// Mitsubishi GX Works2 project: PCL_레더   PLC: Q02/Q02H

PROGRAM MAIN
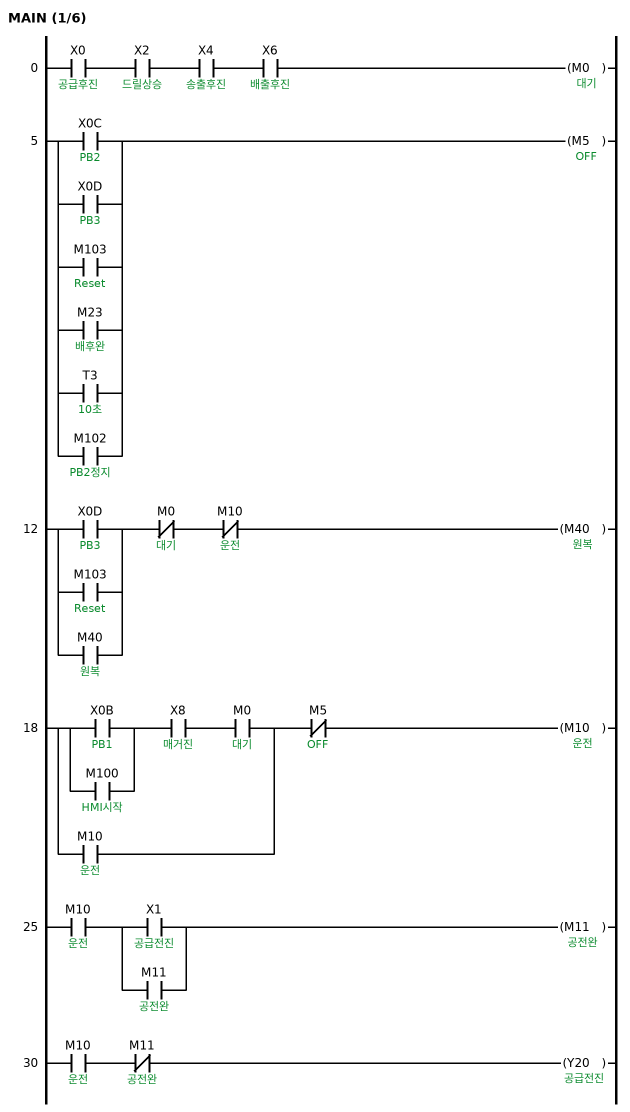
0     LD      X0  ; 공급후진
      AND     X2  ; 드릴상승
      AND     X4  ; 송출후진
      AND     X6  ; 배출후진
      OUT     M0  ; 대기
5     LD      X0C  ; PB2
      OR      X0D  ; PB3
      OR      M103  ; Reset
      OR      M23  ; 배후완
      OR      T3  ; 10초
      OR      M102  ; PB2정지
      OUT     M5  ; OFF
12    LD      X0D  ; PB3
      OR      M103  ; Reset
      OR      M40  ; 원복
      ANI     M0  ; 대기
      ANI     M10  ; 운전
      OUT     M40  ; 원복
18    LD      X0B  ; PB1
      OR      M100  ; HMI시작
      AND     X8  ; 매거진
      AND     M0  ; 대기
      OR      M10  ; 운전
      ANI     M5  ; OFF
      OUT     M10  ; 운전
25    LD      M10  ; 운전
      LD      X1  ; 공급전진
      OR      M11  ; 공전완
      ANB
      OUT     M11  ; 공전완
30    LD      M10  ; 운전
      ANI     M11  ; 공전완
      OUT     Y20  ; 공급전진
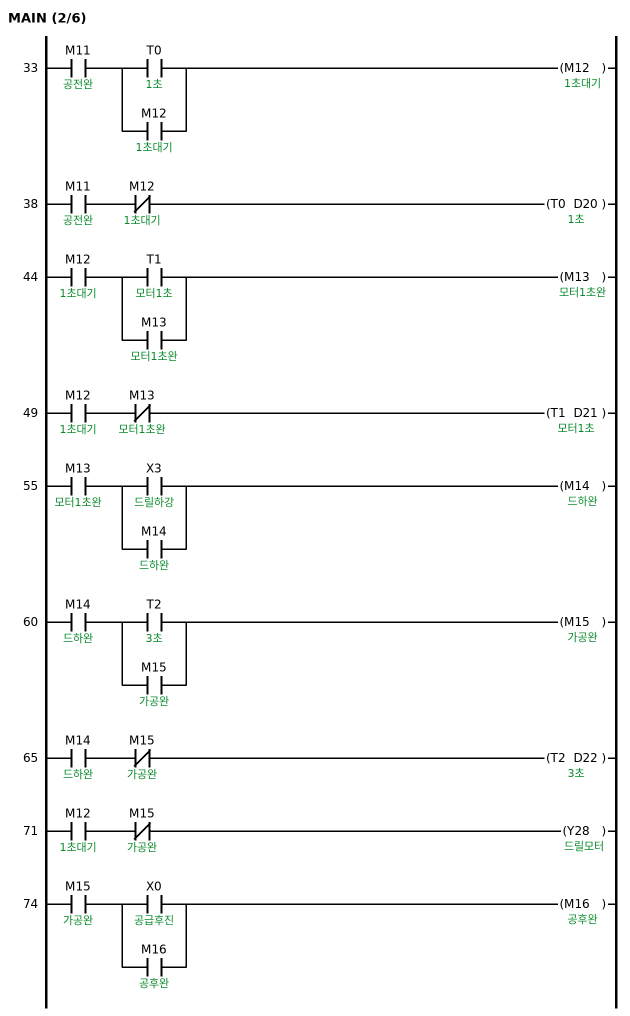
33    LD      M11  ; 공전완
      LD      T0  ; 1초
      OR      M12  ; 1초대기
      ANB
      OUT     M12  ; 1초대기
38    LD      M11  ; 공전완
      ANI     M12  ; 1초대기
      OUT     T0 D20  ; 1초
44    LD      M12  ; 1초대기
      LD      T1  ; 모터1초
      OR      M13  ; 모터1초완
      ANB
      OUT     M13  ; 모터1초완
49    LD      M12  ; 1초대기
      ANI     M13  ; 모터1초완
      OUT     T1 D21  ; 모터1초
55    LD      M13  ; 모터1초완
      LD      X3  ; 드릴하강
      OR      M14  ; 드하완
      ANB
      OUT     M14  ; 드하완
60    LD      M14  ; 드하완
      LD      T2  ; 3초
      OR      M15  ; 가공완
      ANB
      OUT     M15  ; 가공완
65    LD      M14  ; 드하완
      ANI     M15  ; 가공완
      OUT     T2 D22  ; 3초
71    LD      M12  ; 1초대기
      ANI     M15  ; 가공완
      OUT     Y28  ; 드릴모터
74    LD      M15  ; 가공완
      LD      X0  ; 공급후진
      OR      M16  ; 공후완
      ANB
      OUT     M16  ; 공후완
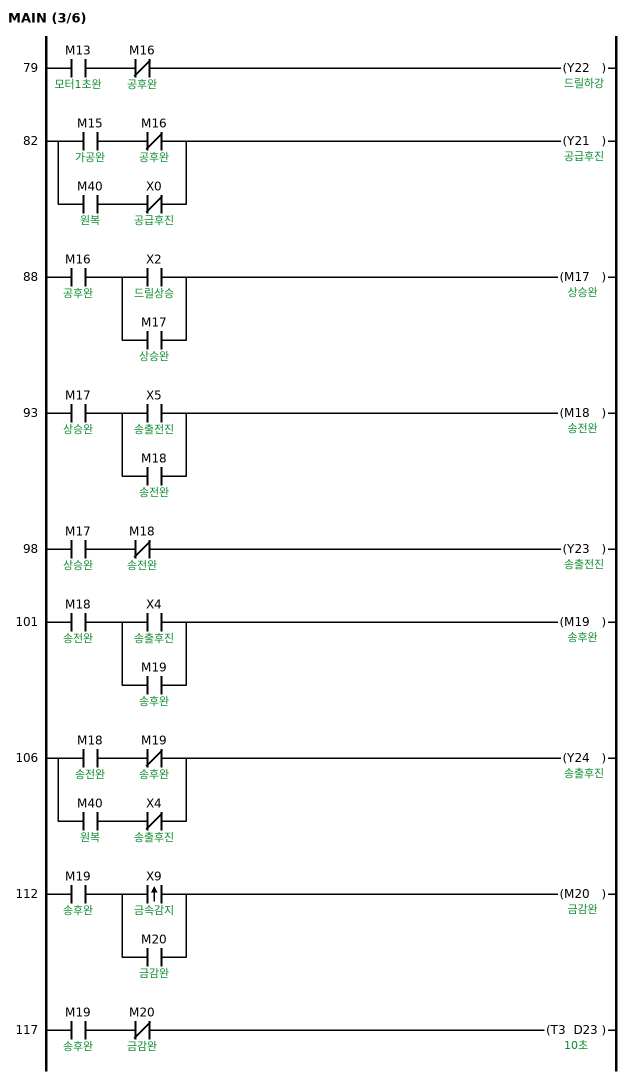
79    LD      M13  ; 모터1초완
      ANI     M16  ; 공후완
      OUT     Y22  ; 드릴하강
82    LD      M15  ; 가공완
      ANI     M16  ; 공후완
      LD      M40  ; 원복
      ANI     X0  ; 공급후진
      ORB
      OUT     Y21  ; 공급후진
88    LD      M16  ; 공후완
      LD      X2  ; 드릴상승
      OR      M17  ; 상승완
      ANB
      OUT     M17  ; 상승완
93    LD      M17  ; 상승완
      LD      X5  ; 송출전진
      OR      M18  ; 송전완
      ANB
      OUT     M18  ; 송전완
98    LD      M17  ; 상승완
      ANI     M18  ; 송전완
      OUT     Y23  ; 송출전진
101   LD      M18  ; 송전완
      LD      X4  ; 송출후진
      OR      M19  ; 송후완
      ANB
      OUT     M19  ; 송후완
106   LD      M18  ; 송전완
      ANI     M19  ; 송후완
      LD      M40  ; 원복
      ANI     X4  ; 송출후진
      ORB
      OUT     Y24  ; 송출후진
112   LD      M19  ; 송후완
      LDP     X9  ; 금속감지
      OR      M20  ; 금감완
      ANB
      OUT     M20  ; 금감완
117   LD      M19  ; 송후완
      ANI     M20  ; 금감완
      OUT     T3 D23  ; 10초
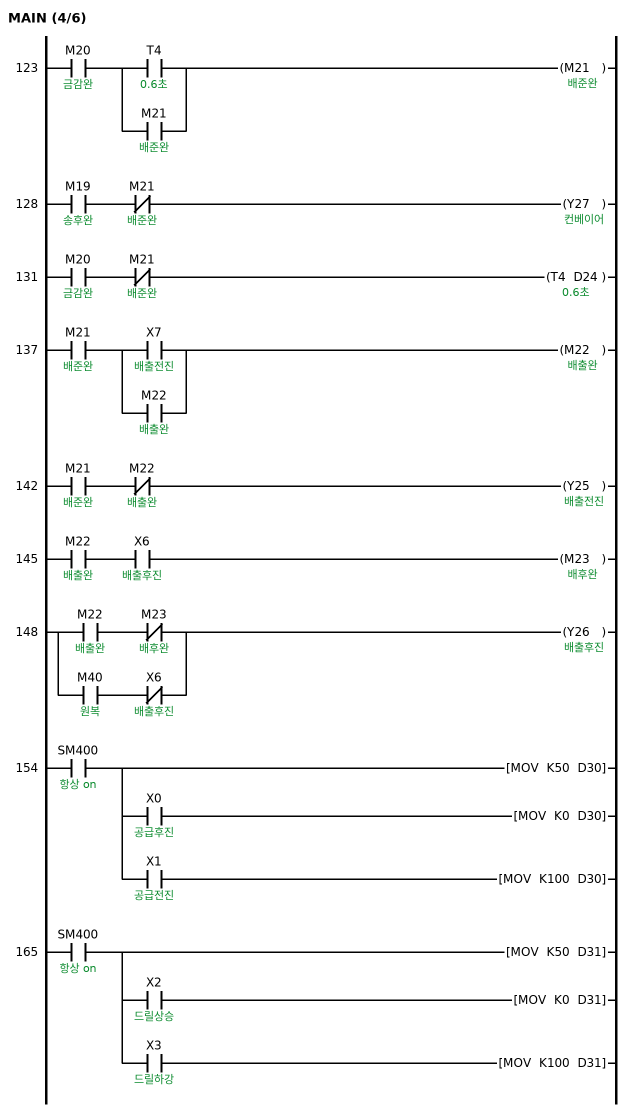
123   LD      M20  ; 금감완
      LD      T4  ; 0.6초
      OR      M21  ; 배준완
      ANB
      OUT     M21  ; 배준완
128   LD      M19  ; 송후완
      ANI     M21  ; 배준완
      OUT     Y27  ; 컨베이어
131   LD      M20  ; 금감완
      ANI     M21  ; 배준완
      OUT     T4 D24  ; 0.6초
137   LD      M21  ; 배준완
      LD      X7  ; 배출전진
      OR      M22  ; 배출완
      ANB
      OUT     M22  ; 배출완
142   LD      M21  ; 배준완
      ANI     M22  ; 배출완
      OUT     Y25  ; 배출전진
145   LD      M22  ; 배출완
      AND     X6  ; 배출후진
      OUT     M23  ; 배후완
148   LD      M22  ; 배출완
      ANI     M23  ; 배후완
      LD      M40  ; 원복
      ANI     X6  ; 배출후진
      ORB
      OUT     Y26  ; 배출후진
154   LD      SM400  ; 항상 on
      MOV     K50 D30
      MPS
      AND     X0  ; 공급후진
      MOV     K0 D30
      MPP
      AND     X1  ; 공급전진
      MOV     K100 D30
165   LD      SM400  ; 항상 on
      MOV     K50 D31
      MPS
      AND     X2  ; 드릴상승
      MOV     K0 D31
      MPP
      AND     X3  ; 드릴하강
      MOV     K100 D31
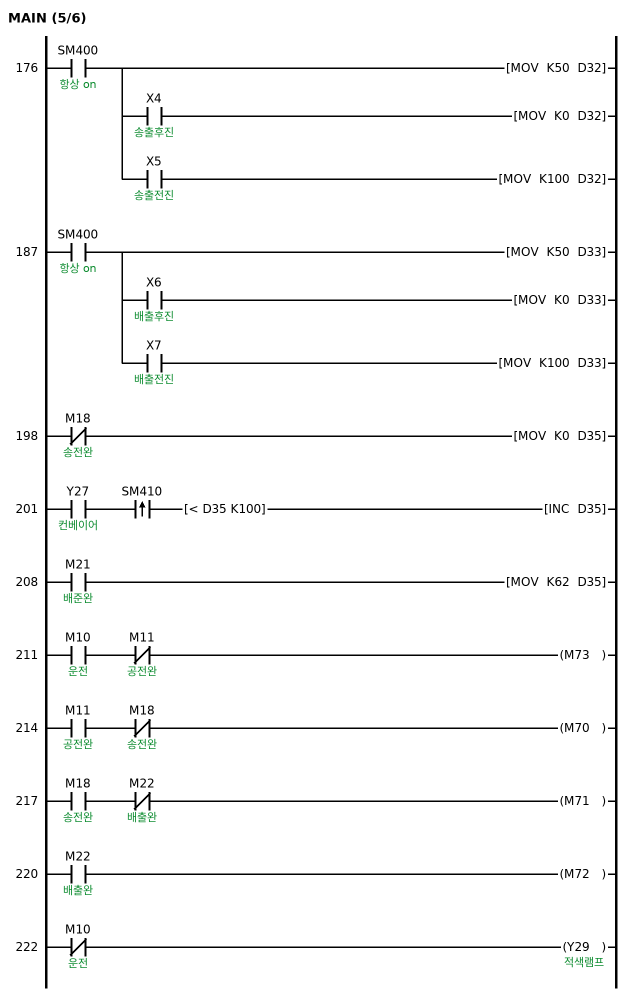
176   LD      SM400  ; 항상 on
      MOV     K50 D32
      MPS
      AND     X4  ; 송출후진
      MOV     K0 D32
      MPP
      AND     X5  ; 송출전진
      MOV     K100 D32
187   LD      SM400  ; 항상 on
      MOV     K50 D33
      MPS
      AND     X6  ; 배출후진
      MOV     K0 D33
      MPP
      AND     X7  ; 배출전진
      MOV     K100 D33
198   LDI     M18  ; 송전완
      MOV     K0 D35
201   LD      Y27  ; 컨베이어
      ANDP    SM410
      AND<    D35 K100
      INC     D35
208   LD      M21  ; 배준완
      MOV     K62 D35
211   LD      M10  ; 운전
      ANI     M11  ; 공전완
      OUT     M73
214   LD      M11  ; 공전완
      ANI     M18  ; 송전완
      OUT     M70
217   LD      M18  ; 송전완
      ANI     M22  ; 배출완
      OUT     M71
220   LD      M22  ; 배출완
      OUT     M72
222   LDI     M10  ; 운전
      OUT     Y29  ; 적색램프
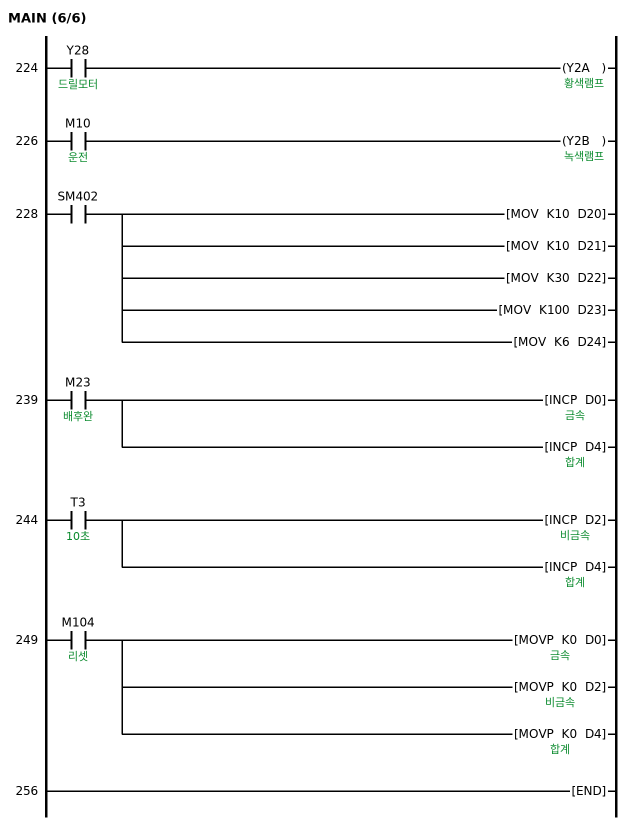
224   LD      Y28  ; 드릴모터
      OUT     Y2A  ; 황색램프
226   LD      M10  ; 운전
      OUT     Y2B  ; 녹색램프
228   LD      SM402
      MOV     K10 D20
      MOV     K10 D21
      MOV     K30 D22
      MOV     K100 D23
      MOV     K6 D24
239   LD      M23  ; 배후완
      INCP    D0  ; 금속
      INCP    D4  ; 합계
244   LD      T3  ; 10초
      INCP    D2  ; 비금속
      INCP    D4
249   LD      M104  ; 리셋
      MOVP    K0 D0
      MOVP    K0 D2
      MOVP    K0 D4
256   END
END_PROGRAM
